Fanuc KAREL source: kd00044.KL

-- PROVISIONAL review KL for V770-1; original PC SHA256 587f4ae1790476c7e5cb29ae4795cda703e4f2176f91f18303fae9b5a44c6ae0
-- Incomplete behavior may be omitted. Consult companion uncertainty JSON. Do not deploy.
PROGRAM KD00044
%NOLOCKGROUP
VAR
  I : INTEGER
  J : INTEGER
  B : BOOLEAN
  R : REAL
  S : STRING[80]
-- UNRESOLVED_DECL G type=00011e
BEGIN
  -- UNRESOLVED_PC offsets 5-12; opcodes 9D,23
  -- UNRESOLVED_PC offsets 17-21; opcodes 7F
END KD00044
